(* Tests LinkFactory and FB_Links: that a link holds copies of the context it points at, that
   the collection owns its links, keeps their order and refuses links beyond its bound.

   Every test releases the contexts and links it builds before returning. *)
FUNCTION_BLOCK FB_TestLinks EXTENDS FB_TestSuite

THIS^.testFromContextCopiesIdentity();
THIS^.testFromContextRejectsInvalidInput();
THIS^.testFromSpanLinksToTheSpan();
THIS^.testPushTakesOwnershipInOrder();
THIS^.testPushRefusesWhenFull();
THIS^.testFromLinkCopiesLink();
THIS^.testFromLinkRejectsInvalidInput();

(* Builds a span context whose identifier bytes are all seed, for a test to link to. *)
METHOD _buildContext
VAR_IN_OUT
	pDest: POINTER TO FB_SpanContext;
END_VAR
VAR_INPUT
	seed: BYTE;
	traceFlags: UDINT;
END_VAR
VAR
	_traceId: FB_TraceId;
	_spanId: FB_SpanId;
END_VAR
MEMSET(ADR(_traceId.bytes), seed, SIZEOF(_traceId.bytes));
MEMSET(ADR(_spanId.bytes), seed, SIZEOF(_spanId.bytes));
ContextFactory.buildContext(
	pDest:=pDest,
	pTraceId:=ADR(_traceId),
	pSpanId:=ADR(_spanId),
	pTraceState:=0,
	traceFlags:=traceFlags
);
END_METHOD

(* A link holds copies of the context's identity and trace state, so it outlives the context.
   Its flags carry the context's trace flags and remoteness. *)
METHOD testFromContextCopiesIdentity : REFERENCE TO FB_Test
VAR
	pContext: POINTER TO FB_SpanContext;
	pLink: POINTER TO FB_Link;
	traceId: FB_TraceId;
	spanId: FB_SpanId;
	traceStateText: T_MaxString := 'vendor=abc';
	pTraceState: POINTER TO FB_TraceState;
	success: BOOL;
	reason: E_LinkFailureReason;
END_VAR
TcUnit.TEST('testFromContextCopiesIdentity');
	MEMSET(ADR(traceId.bytes), 16#AA, SIZEOF(traceId.bytes));
	MEMSET(ADR(spanId.bytes), 16#BB, SIZEOF(spanId.bytes));
	TraceStateFactory.parse(pDest:=pTraceState, pHeader:=ADR(traceStateText));
	ContextFactory.buildContext(
		pDest:=pContext,
		pTraceId:=ADR(traceId),
		pSpanId:=ADR(spanId),
		pTraceState:=pTraceState,
		traceFlags:=16#301  // sampled, remoteness known, remote
	);
	IF pTraceState <> 0 THEN pTraceState^.delete(pSelf:=pTraceState); END_IF

	success := LinkFactory.fromContext(pDest:=pLink, pContext:=pContext, failureReason=>reason);
	THIS^.AssertTrue(success, 'Expected the link to build');
	THIS^.AssertEquals_UDINT(TO_UDINT(E_LinkFailureReason.NA), TO_UDINT(reason), 'Expected no failure reason');

	// the context is borrowed, so it can be released before the link
	IF pContext <> 0 THEN pContext^.delete(pSelf:=pContext); END_IF

	IF pLink <> 0 THEN
		THIS^.AssertTrue(
			pLink^.traceId <> 0 AND_THEN MEMCMP(ADR(pLink^.traceId^.bytes), ADR(traceId.bytes), SIZEOF(traceId.bytes)) = 0,
			'Expected the linked trace id'
		);
		THIS^.AssertTrue(
			pLink^.spanId <> 0 AND_THEN MEMCMP(ADR(pLink^.spanId^.bytes), ADR(spanId.bytes), SIZEOF(spanId.bytes)) = 0,
			'Expected the linked span id'
		);
		THIS^.AssertTrue(pLink^.traceState <> 0, 'Expected the trace state to be copied');
		IF pLink^.traceState <> 0 THEN
			THIS^.AssertEquals_STRING('vendor=abc', pLink^.traceState^.pString^, 'Expected the trace state text');
		END_IF
		THIS^.AssertEquals_UDINT(16#301, pLink^.flags, 'Expected sampled, remoteness known, remote (16#301)');
		THIS^.AssertEquals_UDINT(0, pLink^.attributes.count, 'Expected no attributes');
		pLink^.delete(pSelf:=pLink);
	END_IF
TcUnit.TEST_FINISHED();
END_METHOD

(* fromContext refuses an assigned destination, a null context and an all zero context,
   and allocates nothing when it does. *)
METHOD testFromContextRejectsInvalidInput : REFERENCE TO FB_Test
VAR
	pContext: POINTER TO FB_SpanContext;
	pZero: POINTER TO FB_SpanContext;
	pLink: POINTER TO FB_Link;
	pOther: POINTER TO FB_Link;
	success: BOOL;
	reason: E_LinkFailureReason;
END_VAR
TcUnit.TEST('testFromContextRejectsInvalidInput');
	THIS^._buildContext(pDest:=pContext, seed:=16#11, traceFlags:=16#101);  // sampled, remoteness known, local
	THIS^._buildContext(pDest:=pZero, seed:=0, traceFlags:=0);  // all zero ids: an invalid context

	success := LinkFactory.fromContext(pDest:=pLink, pContext:=0, failureReason=>reason);
	THIS^.AssertFalse(success, 'Expected a null context to be refused');
	THIS^.AssertEquals_UDINT(TO_UDINT(E_LinkFailureReason.CONTEXT_POINTER_NULL), TO_UDINT(reason), 'Expected CONTEXT_POINTER_NULL');
	THIS^.AssertTrue(pLink = 0, 'Expected nothing to be allocated for a null context');

	success := LinkFactory.fromContext(pDest:=pLink, pContext:=pZero, failureReason=>reason);
	THIS^.AssertFalse(success, 'Expected an invalid context to be refused');
	THIS^.AssertEquals_UDINT(TO_UDINT(E_LinkFailureReason.CONTEXT_INVALID), TO_UDINT(reason), 'Expected CONTEXT_INVALID');
	THIS^.AssertTrue(pLink = 0, 'Expected nothing to be allocated for an invalid context');

	LinkFactory.fromContext(pDest:=pLink, pContext:=pContext);
	pOther := pLink;
	success := LinkFactory.fromContext(pDest:=pLink, pContext:=pContext, failureReason=>reason);
	THIS^.AssertFalse(success, 'Expected an assigned destination to be refused');
	THIS^.AssertEquals_UDINT(TO_UDINT(E_LinkFailureReason.DESTINATION_ALREADY_ASSIGNED), TO_UDINT(reason), 'Expected DESTINATION_ALREADY_ASSIGNED');
	THIS^.AssertTrue(pLink = pOther, 'Expected the destination to be left alone');

	IF pLink <> 0 THEN pLink^.delete(pSelf:=pLink); END_IF
	IF pContext <> 0 THEN pContext^.delete(pSelf:=pContext); END_IF
	IF pZero <> 0 THEN pZero^.delete(pSelf:=pZero); END_IF
TcUnit.TEST_FINISHED();
END_METHOD

(* A link built from a span points at that span, and is local: remoteness is known and not
   remote. A null span is refused. *)
METHOD testFromSpanLinksToTheSpan : REFERENCE TO FB_Test
VAR
	resource: FB_Resource('');
	idGenerator: FB_MockIdGenerator;
	provider: FB_TracerProvider(resource:=resource, idGenerator:=idGenerator, sampler:=TcOtlp_GVL.defaultSampler);
	scope: FB_InstrumentationScope('tracer.test', '1.0.0', '');
	tracer: FB_Tracer(scope:=scope, provider:=provider);
	pSpan: POINTER TO FB_Span;
	pLink: POINTER TO FB_Link;
	success: BOOL;
	reason: E_LinkFailureReason;
END_VAR
TcUnit.TEST('testFromSpanLinksToTheSpan');
	tracer.startSpan(name:='trigger').build(pDest:=pSpan);
	THIS^.AssertTrue(pSpan <> 0, 'Expected the span to build');

	success := LinkFactory.fromSpan(pDest:=pLink, pSpan:=0, failureReason=>reason);
	THIS^.AssertFalse(success, 'Expected a null span to be refused');
	THIS^.AssertEquals_UDINT(TO_UDINT(E_LinkFailureReason.SPAN_POINTER_NULL), TO_UDINT(reason), 'Expected SPAN_POINTER_NULL');

	success := LinkFactory.fromSpan(pDest:=pLink, pSpan:=pSpan, failureReason=>reason);
	THIS^.AssertTrue(success, 'Expected the link to build');
	THIS^.AssertEquals_UDINT(TO_UDINT(E_LinkFailureReason.NA), TO_UDINT(reason), 'Expected no failure reason');
	IF pLink <> 0 AND pSpan <> 0 THEN
		THIS^.AssertTrue(
			MEMCMP(ADR(pLink^.traceId^.bytes), ADR(pSpan^.traceId^.bytes), SIZEOF(pSpan^.traceId^.bytes)) = 0,
			'Expected the span$'s trace id'
		);
		THIS^.AssertTrue(
			MEMCMP(ADR(pLink^.spanId^.bytes), ADR(pSpan^.spanId^.bytes), SIZEOF(pSpan^.spanId^.bytes)) = 0,
			'Expected the span$'s span id'
		);
		THIS^.AssertEquals_UDINT(16#101, pLink^.flags, 'Expected the sampled bit and a known local context (16#101)');
	END_IF

	IF pLink <> 0 THEN pLink^.delete(pSelf:=pLink); END_IF
	IF pSpan <> 0 THEN pSpan^.delete(pSelf:=pSpan); END_IF
TcUnit.TEST_FINISHED();
END_METHOD

(* push takes ownership and clears the caller's pointer; next walks the links oldest first
   without taking them, and pop hands them back in the same order. *)
METHOD testPushTakesOwnershipInOrder : REFERENCE TO FB_Test
VAR
	links: FB_Links(maxCount:=TcOtlp_GVL.DEFAULT_MAX_LINK_COUNT);
	pFirst: POINTER TO FB_SpanContext;
	pSecond: POINTER TO FB_SpanContext;
	pLink: POINTER TO FB_Link;
	pWalked: POINTER TO FB_Link;
	success: BOOL;
	reason: E_LinkFailureReason;
END_VAR
TcUnit.TEST('testPushTakesOwnershipInOrder');
	// 16#101: sampled, remoteness known, local; the seed byte tells the links apart
	THIS^._buildContext(pDest:=pFirst, seed:=16#11, traceFlags:=16#101);
	THIS^._buildContext(pDest:=pSecond, seed:=16#22, traceFlags:=16#101);

	LinkFactory.fromContext(pDest:=pLink, pContext:=pFirst);
	success := links.push(pValue:=pLink, failureReason=>reason);
	THIS^.AssertTrue(success, 'Expected the first push to succeed');
	THIS^.AssertEquals_UDINT(TO_UDINT(E_LinkFailureReason.NA), TO_UDINT(reason), 'Expected no failure reason');
	THIS^.AssertTrue(pLink = 0, 'Expected push to clear the caller$'s pointer');
	LinkFactory.fromContext(pDest:=pLink, pContext:=pSecond);
	links.push(pValue:=pLink);
	THIS^.AssertEquals_UDINT(2, links.count, 'Expected two links');

	links.reset();
	pWalked := links.next();
	THIS^.AssertTrue(pWalked <> 0 AND_THEN pWalked^.spanId^.bytes[0] = 16#11, 'Expected next to start at the oldest link');
	pWalked := links.next();
	THIS^.AssertTrue(pWalked <> 0 AND_THEN pWalked^.spanId^.bytes[0] = 16#22, 'Expected next to reach the second link');
	THIS^.AssertTrue(links.next() = 0, 'Expected next to end after the last link');
	THIS^.AssertEquals_UDINT(2, links.count, 'Expected walking to leave the links in place');

	success := links.pop(pValue:=pLink, failureReason=>reason);
	THIS^.AssertTrue(success AND_THEN pLink^.spanId^.bytes[0] = 16#11, 'Expected pop to return the oldest link');
	success := links.pop(pValue:=pLink, failureReason=>reason);
	THIS^.AssertFalse(success, 'Expected pop into an assigned destination to fail');
	THIS^.AssertEquals_UDINT(TO_UDINT(E_LinkFailureReason.DESTINATION_ALREADY_ASSIGNED), TO_UDINT(reason), 'Expected DESTINATION_ALREADY_ASSIGNED');
	IF pLink <> 0 THEN pLink^.delete(pSelf:=pLink); END_IF

	links.pop(pValue:=pLink);
	IF pLink <> 0 THEN pLink^.delete(pSelf:=pLink); END_IF
	success := links.pop(pValue:=pLink, failureReason=>reason);
	THIS^.AssertFalse(success, 'Expected pop from an empty collection to fail');
	THIS^.AssertEquals_UDINT(TO_UDINT(E_LinkFailureReason.LINKS_EMPTY), TO_UDINT(reason), 'Expected LINKS_EMPTY');
	THIS^.AssertEquals_UDINT(0, links.count, 'Expected no links left');

	IF pFirst <> 0 THEN pFirst^.delete(pSelf:=pFirst); END_IF
	IF pSecond <> 0 THEN pSecond^.delete(pSelf:=pSecond); END_IF
TcUnit.TEST_FINISHED();
END_METHOD

(* A full collection keeps its links and refuses the new one: the caller keeps it, and it is
   counted as dropped. A null link is refused without being counted. free releases every link. *)
METHOD testPushRefusesWhenFull : REFERENCE TO FB_Test
VAR
	links: FB_Links(maxCount:=1);
	pContext: POINTER TO FB_SpanContext;
	pLink: POINTER TO FB_Link;
	pRefused: POINTER TO FB_Link;
	success: BOOL;
	reason: E_LinkFailureReason;
END_VAR
TcUnit.TEST('testPushRefusesWhenFull');
	THIS^._buildContext(pDest:=pContext, seed:=16#11, traceFlags:=16#101);  // sampled, remoteness known, local

	success := links.push(pValue:=pLink, failureReason=>reason);
	THIS^.AssertFalse(success, 'Expected a null link to be refused');
	THIS^.AssertEquals_UDINT(TO_UDINT(E_LinkFailureReason.LINK_POINTER_NULL), TO_UDINT(reason), 'Expected LINK_POINTER_NULL');

	LinkFactory.fromContext(pDest:=pLink, pContext:=pContext);
	links.push(pValue:=pLink);
	LinkFactory.fromContext(pDest:=pLink, pContext:=pContext);
	pRefused := pLink;
	success := links.push(pValue:=pLink, failureReason=>reason);
	THIS^.AssertFalse(success, 'Expected a push beyond maxCount to fail');
	THIS^.AssertEquals_UDINT(TO_UDINT(E_LinkFailureReason.LINK_COUNT_LIMIT_REACHED), TO_UDINT(reason), 'Expected LINK_COUNT_LIMIT_REACHED');
	THIS^.AssertTrue(pLink = pRefused, 'Expected the caller to keep the refused link');
	THIS^.AssertEquals_UDINT(1, links.count, 'Expected the first link to be kept');
	THIS^.AssertEquals_UDINT(1, links.droppedCount, 'Expected the refused link to be counted');
	IF pLink <> 0 THEN pLink^.delete(pSelf:=pLink); END_IF

	THIS^.AssertTrue(links.free(), 'Expected free to release every link');
	THIS^.AssertEquals_UDINT(0, links.count, 'Expected no links after free');
	THIS^.AssertEquals_UDINT(0, links.droppedCount, 'Expected free to clear droppedCount');

	IF pContext <> 0 THEN pContext^.delete(pSelf:=pContext); END_IF
TcUnit.TEST_FINISHED();
END_METHOD

(* fromLink gives the copy its own identity, trace state and attributes. *)
METHOD testFromLinkCopiesLink : REFERENCE TO FB_Test
VAR
	pContext: POINTER TO FB_SpanContext;
	pLink: POINTER TO FB_Link;
	pCopy: POINTER TO FB_Link;
	reason: E_LinkFailureReason;
END_VAR
TcUnit.TEST('testFromLinkCopiesLink');
	THIS^._buildContext(pDest:=pContext, seed:=5, traceFlags:=1);  // sampled only
	LinkFactory.fromContext(pDest:=pLink, pContext:=pContext, failureReason=>reason);
	THIS^.AssertTrue(pLink <> 0, 'Expected the source link to build');
	IF pLink <> 0 THEN
		pLink^.attributes.setStringAttribute('k', 'v');
		THIS^.AssertTrue(LinkFactory.fromLink(pDest:=pCopy, pSrc:=pLink, failureReason=>reason), 'Expected fromLink to succeed');
		IF pCopy <> 0 THEN
			THIS^.AssertTrue(pCopy^.traceId <> 0 AND_THEN pCopy^.traceId <> pLink^.traceId, 'Expected a copied trace id');
			THIS^.AssertTrue(pCopy^.spanId <> 0 AND_THEN pCopy^.spanId <> pLink^.spanId, 'Expected a copied span id');
			THIS^.AssertEquals_UDINT(pLink^.flags, pCopy^.flags, 'Expected the flags');
			THIS^.AssertEquals_UDINT(1, pCopy^.attributes.count, 'Expected the attribute');
			pLink^.delete(pSelf:=pLink);
			THIS^.AssertTrue(pCopy^.traceId^.bytes[0] = 5 AND pCopy^.spanId^.bytes[0] = 5, 'Expected the identity to outlive the source');
			pCopy^.delete(pSelf:=pCopy);
		END_IF
		IF pLink <> 0 THEN pLink^.delete(pSelf:=pLink); END_IF
	END_IF
	IF pContext <> 0 THEN pContext^.delete(pSelf:=pContext); END_IF
TcUnit.TEST_FINISHED();
END_METHOD

(* fromLink refuses a missing source and an assigned destination. *)
METHOD testFromLinkRejectsInvalidInput : REFERENCE TO FB_Test
VAR
	pLink: POINTER TO FB_Link;
	pDest: POINTER TO FB_Link;
	reason: E_LinkFailureReason;
END_VAR
TcUnit.TEST('testFromLinkRejectsInvalidInput');
	THIS^.AssertFalse(LinkFactory.fromLink(pDest:=pDest, pSrc:=0, failureReason=>reason), 'Expected a null source to fail');
	THIS^.AssertEquals_UDINT(TO_UDINT(E_LinkFailureReason.LINK_POINTER_NULL), TO_UDINT(reason), 'Expected LINK_POINTER_NULL');

	pLink := __NEW(FB_Link);  // built by hand: LinkFactory refuses a link with no identity
	THIS^.AssertFalse(LinkFactory.fromLink(pDest:=pDest, pSrc:=pLink, failureReason=>reason), 'Expected an empty link to fail');
	THIS^.AssertEquals_UDINT(TO_UDINT(E_LinkFailureReason.CONTEXT_INVALID), TO_UDINT(reason), 'Expected CONTEXT_INVALID');

	pDest := pLink;
	THIS^.AssertFalse(LinkFactory.fromLink(pDest:=pDest, pSrc:=pLink, failureReason=>reason), 'Expected an assigned destination to fail');
	THIS^.AssertEquals_UDINT(
		TO_UDINT(E_LinkFailureReason.DESTINATION_ALREADY_ASSIGNED),
		TO_UDINT(reason),
		'Expected DESTINATION_ALREADY_ASSIGNED'
	);
	THIS^.AssertTrue(pDest = pLink, 'Expected the destination to be left alone');
	IF pLink <> 0 THEN pLink^.delete(pSelf:=pLink); END_IF
TcUnit.TEST_FINISHED();
END_METHOD

END_FUNCTION_BLOCK

(* stored: Version 1.1.0.1
   POU FB_TestLinks: Id {774cbd45-c83b-4748-9cdc-bfbacf04f1cc}, SpecialFunc None
   Method _buildContext: Id {cc0180b8-bb00-4066-86bc-df7b7037186f}
   Method testFromContextCopiesIdentity: Id {204ccd02-c522-40e9-b35f-c11b0f7f8727}
   Method testFromContextRejectsInvalidInput: Id {22ab2495-4520-4a85-b906-bbfa89e9ea0a}
   Method testFromSpanLinksToTheSpan: Id {fa2845c8-83a6-46af-a075-0e77a5da39b9}
   Method testPushTakesOwnershipInOrder: Id {a1d4c8f6-7340-4c6d-9461-226f7c917ddf}
   Method testPushRefusesWhenFull: Id {25eef890-4e51-4894-8fce-f5ac86e0c639}
   Method testFromLinkCopiesLink: Id {bb2598d0-ced5-42be-b32d-b2a360498f53}
   Method testFromLinkRejectsInvalidInput: Id {a95df6e9-e0a0-4d27-a0f5-7ad4eb6fcc06} *)
